(* IEC 61131-3 sources: plc-vscode/tests/st/all/rusty/tests/lit/multi/header_generator/number_container, 1 file *)

(* ---- number_container_prog.st ---- *)
FUNCTION main
VAR
    numberContainerFb : NumberContainer;
END_VAR
    numberContainerFb();
    PrintNumber(numberContainerFb.GetMemberValue());  // CHECK: The number you asked for: 42
END_FUNCTION
